Fanuc KAREL source: KC00031.KL

PROGRAM KC00031
%NOLOCKGROUP
%ENVIRONMENT TIM
VAR
  I: INTEGER
  J: INTEGER
  K: INTEGER
  R: REAL
  B: BOOLEAN
  S: STRING[80]
  T: STRING[80]
  P: PATH
  Q: PATH
  AI: ARRAY[8] OF INTEGER
  AB: ARRAY[244] OF BYTE
BEGIN
  I = GET_USEC_SUB(J,K)
END KC00031
